Fanuc KAREL source: KT00937.KL

PROGRAM KT00937
%NOLOCKGROUP
VAR
  ENTRY: INTEGER
  PNAME: STRING[80]
  VNAME: STRING[80]
  STATUS: INTEGER
  VALUE: ARRAY[2] OF BYTE
BEGIN
  ENTRY = 0
  PNAME = ''
  VNAME = 'VALUE'
  VALUE[1] = 2
  GET_VAR(ENTRY, PNAME, VNAME, VALUE[1], STATUS)
END KT00937
